// TIA Portal V20 export
VAR_GLOBAL   // PLC tag table "LASER_IN_datalogic"
   LASER_OFF AT %I400.0 : Bool;
   LASER_WARM_UP AT %I400.1 : Bool;
   LASER_WAIT_FOR_START AT %I400.2 : Bool;
   LASER_STANDBY AT %I400.3 : Bool;
   LASER_STANDBY_SHUTTER_CLOSED AT %I400.4 : Bool;
   LASER_READY AT %I400.5 : Bool;
   LASER_EMISSION AT %I400.6 : Bool;
   LASER_BUSSY_SHUTTER_CLOSED AT %I401.0 : Bool;
   LASER_WARNING AT %I401.1 : Bool;
   LASER_ERROR AT %I401.2 : Bool;
   COMMAND_EXECUTING AT %I402.0 : Bool;
   COMMAND_ERROR AT %I402.1 : Bool;
   PROTOCOL_ERROR AT %I402.2 : Bool;
   PROTOCOL_BOOT_UP AT %I403.7 : Bool;
   COMMAND_ERROR_CODE AT %IB404 : Byte;
   PROTOCOL_ERROR_CODE AT %IB405 : Byte;
   RESERVE_I_6_BYTE AT %IB406 : Byte;
   RESERVE_I_7_BYTE AT %IB407 : Byte;
   RESERVE_I_8_BYTE AT %IB408 : Byte;
   RESERVE_I_9_BYTE AT %IB409 : Byte;
   START_MARKING_IN AT %I410.0 : Bool;
   STOP_SYSTEM_IN AT %I410.1 : Bool;
   GET_PNIO_PROTOCOL_VERSION_IN AT %I411.0 : Bool;
   GET_LASER_ENGINE_VERSION AT %I411.1 : Bool;
   OPEN_DOCUMENT_FROM_DEVICE AT %I412.0 : Bool;
   SAVE_DOCUMENT AT %I412.1 : Bool;
   GET_DATA_FIELD_VALUE_IN AT %I412.2 : Bool;
   SET_DATA_FIELD_VALUE_IN AT %I412.3 : Bool;
   GET_GLOBAL_COUNTER_VALUE_IN AT %I412.4 : Bool;
   SET_GLOBAL_COUNTER_VALUE_IN AT %I412.5 : Bool;
   GET_GLOBAL_STRING_VALUE_IN AT %I412.6 : Bool;
   SET_GLOBAL_STRING_VALUE_IN AT %I412.7 : Bool;
   ENABLE_DATA_FIELD_IN AT %I413.0 : Bool;
   DISABLE_DATA_FIELD_IN AT %I413.1 : Bool;
   MOVE_END_ROTATE_DOCUMENT AT %I414.0 : Bool;
   MOVE_DATA_FIELD_IN AT %I414.1 : Bool;
   RESERVE_I_15_BYTE AT %IB415 : Byte;
   RESERVE_I_16_BYTE AT %IB416 : Byte;
   RESERVE_I_17_BYTE AT %IB417 : Byte;
   MOVE_AXIS_IN AT %I418.0 : Bool;
   RESET_AXIS_IN AT %I418.1 : Bool;
   STOP_AXIS_IN AT %I418.2 : Bool;
   START_AUTOFOCUS_IN AT %I418.3 : Bool;
   STOP_AUTOFOCUS_IN AT %I418.4 : Bool;
   SET_FOCUS_DISTANCE_REFERENCE_IN AT %I418.5 : Bool;
   RESERVE_I_19_BYTE AT %IB419 : Byte;
   X_AXIS_ENABLED AT %I420.0 : Bool;
   Y_AXIS_ENABLED AT %I420.1 : Bool;
   Z_AXIS_ENABLED AT %I420.2 : Bool;
   R_AXIS_ENABLED AT %I420.3 : Bool;
   X_AXIS_HOME AT %I420.4 : Bool;
   Y_AXIS_HOME AT %I420.5 : Bool;
   Z_AXIS_HOME AT %I420.6 : Bool;
   R_AXIS_HOME AT %I420.7 : Bool;
   X_AXIS_MOVEMENT AT %I421.0 : Bool;
   Y_AXIS_MOVEMENT AT %I421.1 : Bool;
   Z_AXIS_MOVEMENT AT %I421.2 : Bool;
   R_AXIS_MOVEMENT AT %I421.3 : Bool;
   Z_ASIS_IN_ON_FOCUS AT %I421.4 : Bool;
   FOCUS_DISTANCE_SENSOR_IS_AVAILABLE AT %I421.5 : Bool;
   RESERVE_I_22_BYTE AT %IB422 : Byte;
   RESERVE_I_23_BYTE AT %IB423 : Byte;
   SET_OUTPUT AT %I424.0 : Bool;
   RESET_OUTPUT_IN AT %I424.1 : Bool;
   RRESERVE_I_25_BYTE AT %IB425 : Byte;
   I_O_PORT_LASER_OUTPUT_STATUS_0 AT %I426.0 : Bool;
   I_O_PORT_LASER_OUTPUT_STATUS_1 AT %I426.1 : Bool;
   I_O_PORT_LASER_OUTPUT_STATUS_2 AT %I426.2 : Bool;
   I_O_PORT_LASER_OUTPUT_STATUS_3 AT %I426.3 : Bool;
   I_O_PORT_LASER_OUTPUT_STATUS_4 AT %I426.4 : Bool;
   I_O_PORT_LASER_OUTPUT_STATUS_5 AT %I426.5 : Bool;
   I_O_PORT_LASER_OUTPUT_STATUS_6 AT %I426.6 : Bool;
   I_O_PORT_LASER_OUTPUT_STATUS_7 AT %I426.7 : Bool;
   I_O_PORT_LASER_OUTPUT_STATUS_8 AT %I427.0 : Bool;
   I_O_PORT_LASER_OUTPUT_STATUS_9 AT %I427.1 : Bool;
   I_O_PORT_LASER_OUTPUT_STATUS_10 AT %I427.2 : Bool;
   I_O_PORT_LASER_OUTPUT_STATUS_11 AT %I427.3 : Bool;
   I_O_PORT_LASER_OUTPUT_STATUS_12 AT %I427.4 : Bool;
   I_O_PORT_LASER_OUTPUT_STATUS_13 AT %I427.5 : Bool;
   I_O_PORT_LASER_OUTPUT_STATUS_14 AT %I427.6 : Bool;
   I_O_PORT_LASER_OUTPUT_STATUS_15 AT %I427.7 : Bool;
   I_O_PORT_LASER_INPUT_STATUS_0 AT %I428.0 : Bool;
   I_O_PORT_LASER_INPUT_STATUS_1 AT %I428.1 : Bool;
   I_O_PORT_LASER_INPUT_STATUS_2 AT %I428.2 : Bool;
   I_O_PORT_LASER_INPUT_STATUS_3 AT %I428.3 : Bool;
   I_O_PORT_LASER_INPUT_STATUS_4 AT %I428.4 : Bool;
   I_O_PORT_LASER_INPUT_STATUS_5 AT %I428.5 : Bool;
   I_O_PORT_LASER_INPUT_STATUS_6 AT %I428.6 : Bool;
   I_O_PORT_LASER_INPUT_STATUS_7 AT %I428.7 : Bool;
   I_O_PORT_LASER_INPUT_STATUS_8 AT %I429.0 : Bool;
   I_O_PORT_LASER_INPUT_STATUS_9 AT %I429.1 : Bool;
   I_O_PORT_LASER_INPUT_STATUS_10 AT %I429.2 : Bool;
   I_O_PORT_LASER_INPUT_STATUS_11 AT %I429.3 : Bool;
   I_O_PORT_LASER_INPUT_STATUS_12 AT %I429.4 : Bool;
   I_O_PORT_LASER_INPUT_STATUS_13 AT %I429.5 : Bool;
   I_O_PORT_LASER_INPUT_STATUS_14 AT %I429.6 : Bool;
   I_O_PORT_LASER_INPUT_STATUS_15 AT %I429.7 : Bool;
   RESERVE_I_30_BYTE AT %IB430 : Byte;
   RESERVE_I_31_BYTE AT %IB431 : Byte;
   RESERVE_I_32_BYTE AT %IB432 : Byte;
   RESERVE_I_33_BYTE AT %IB433 : Byte;
   GET_ID_MATCH_RESULT_IN AT %I434.1 : Bool;
   GET_ID_MARVIS_CONFIGURATION_IN AT %I434.2 : Bool;
   SET_ID_MARVIS_CONFIGURATION_IN AT %I434.3 : Bool;
   GET_ID_MARVIS_RESULT_IN AT %I434.4 : Bool;
   RESERVE_I_35_BYTE AT %IB435 : Byte;
   MARVIS_RESULT_OK AT %I436.0 : Bool;
   MARVIS_RESULT_FAIL AT %I436.1 : Bool;
   SYMBOL_READ_OK AT %I436.2 : Bool;
   SYMBOL_READ_FAIL AT %I436.3 : Bool;
   SYMBOL_GRADE_RESULT_OK AT %I436.4 : Bool;
   SYMBOL_GRADE_RESULT_FAIL AT %I436.5 : Bool;
   SYMBOL_MATCH_RESULT_OK AT %I436.6 : Bool;
   SYMBOL_MATCH_RESULT_FAIL AT %I436.7 : Bool;
   RESERVE_I_37_BYTE AT %IB437 : Byte;
   READER_STATUS_AVAILABLE AT %I438.1 : Bool;
   READER_STATUS_BZSY AT %I438.2 : Bool;
   READER_STATUS_WARNING AT %I438.3 : Bool;
   READER_STATUS_ERROR AT %I438.4 : Bool;
   RESERVE_I_39_BYTE AT %IB439 : Byte;
   RESERVE_I_40_BYTE AT %IB440 : Byte;
   RESERVE_I_41_BYTE AT %IB441 : Byte;
   RESERVE_I_42_BYTE AT %IB442 : Byte;
   RESERVE_I_43_BYTE AT %IB443 : Byte;
   RESERVE_I_44_BYTE AT %IB444 : Byte;
   RESERVE_I_45_BYTE AT %IB445 : Byte;
   RESERVE_I_46_BYTE AT %IB446 : Byte;
   RESERVE_I_47_BYTE AT %IB447 : Byte;
   RESERVE_I_48_BYTE AT %IB448 : Byte;
   RESERVE_I_49_BYTE AT %IB449 : Byte;
   RESERVE_I_50_BYTE AT %IB450 : Byte;
   RESERVE_I_51_BYTE AT %IB451 : Byte;
   RESERVE_I_52_BYTE AT %IB452 : Byte;
   RESERVE_I_53_BYTE AT %IB453 : Byte;
   RESPONSE_DATE_SIZE AT %IB454 : Byte;
   RESERVE_I_55_BYTE AT %IB455 : Byte;
   RESPONSE_DATA_FIELD_0 AT %IB456 : Byte;
   RESPONSE_DATA_FIELD_1 AT %IB457 : Byte;
   RESPONSE_DATA_FIELD_2 AT %IB458 : Byte;
   RESPONSE_DATA_FIELD_3 AT %IB459 : Byte;
   RESPONSE_DATA_FIELD_4 AT %IB460 : Byte;
   RESPONSE_DATA_FIELD_5 AT %IB461 : Byte;
   RESPONSE_DATA_FIELD_6 AT %IB462 : Byte;
   RESPONSE_DATA_FIELD_7 AT %IB463 : Byte;
   RESPONSE_DATA_FIELD_8 AT %IB464 : Byte;
   RESPONSE_DATA_FIELD_9 AT %IB465 : Byte;
   RESPONSE_DATA_FIELD_10 AT %IB466 : Byte;
   RESPONSE_DATA_FIELD_11 AT %IB467 : Byte;
   RESPONSE_DATA_FIELD_12 AT %IB468 : Byte;
   RESPONSE_DATA_FIELD_13 AT %IB469 : Byte;
   RESPONSE_DATA_FIELD_14 AT %IB470 : Byte;
   RESPONSE_DATA_FIELD_15 AT %IB471 : Byte;
   RESPONSE_DATA_FIELD_16 AT %IB472 : Byte;
   RESPONSE_DATA_FIELD_17 AT %IB473 : Byte;
   RESPONSE_DATA_FIELD_18 AT %IB474 : Byte;
   RESPONSE_DATA_FIELD_19 AT %IB475 : Byte;
   RESPONSE_DATA_FIELD_20 AT %IB476 : Byte;
   RESPONSE_DATA_FIELD_21 AT %IB477 : Byte;
   RESPONSE_DATA_FIELD_22 AT %IB478 : Byte;
   RESPONSE_DATA_FIELD_23 AT %IB479 : Byte;
   RESPONSE_DATA_FIELD_24 AT %IB480 : Byte;
   RESPONSE_DATA_FIELD_25 AT %IB481 : Byte;
   RESPONSE_DATA_FIELD_26 AT %IB482 : Byte;
   RESPONSE_DATA_FIELD_27 AT %IB483 : Byte;
   RESPONSE_DATA_FIELD_28 AT %IB484 : Byte;
   RESPONSE_DATA_FIELD_29 AT %IB485 : Byte;
   RESPONSE_DATA_FIELD_30 AT %IB486 : Byte;
   RESPONSE_DATA_FIELD_31 AT %IB487 : Byte;
   RESPONSE_DATA_FIELD_32 AT %IB488 : Byte;
   RESPONSE_DATA_FIELD_33 AT %IB489 : Byte;
   RESPONSE_DATA_FIELD_34 AT %IB490 : Byte;
   RESPONSE_DATA_FIELD_35 AT %IB491 : Byte;
   RESPONSE_DATA_FIELD_36 AT %IB492 : Byte;
   RESPONSE_DATA_FIELD_37 AT %IB493 : Byte;
   RESPONSE_DATA_FIELD_38 AT %IB494 : Byte;
   RESPONSE_DATA_FIELD_39 AT %IB495 : Byte;
   RESPONSE_DATA_FIELD_40 AT %IB496 : Byte;
   RESPONSE_DATA_FIELD_41 AT %IB497 : Byte;
   RESPONSE_DATA_FIELD_42 AT %IB498 : Byte;
   RESPONSE_DATA_FIELD_43 AT %IB499 : Byte;
   RESPONSE_DATA_FIELD_44 AT %IB500 : Byte;
   RESPONSE_DATA_FIELD_45 AT %IB501 : Byte;
   RESPONSE_DATA_FIELD_46 AT %IB502 : Byte;
   RESPONSE_DATA_FIELD_47 AT %IB503 : Byte;
   RESPONSE_DATA_FIELD_48 AT %IB504 : Byte;
   RESPONSE_DATA_FIELD_49 AT %IB505 : Byte;
   RESPONSE_DATA_FIELD_50 AT %IB506 : Byte;
   RESPONSE_DATA_FIELD_51 AT %IB507 : Byte;
   RESPONSE_DATA_FIELD_52 AT %IB508 : Byte;
   RESPONSE_DATA_FIELD_53 AT %IB509 : Byte;
   RESPONSE_DATA_FIELD_54 AT %IB510 : Byte;
   RESPONSE_DATA_FIELD_55 AT %IB511 : Byte;
   RESPONSE_DATA_FIELD_56 AT %IB512 : Byte;
   RESPONSE_DATA_FIELD_57 AT %IB513 : Byte;
   RESPONSE_DATA_FIELD_58 AT %IB514 : Byte;
   RESPONSE_DATA_FIELD_59 AT %IB515 : Byte;
   RESPONSE_DATA_FIELD_60 AT %IB516 : Byte;
   RESPONSE_DATA_FIELD_61 AT %IB517 : Byte;
   RESPONSE_DATA_FIELD_62 AT %IB518 : Byte;
   RESPONSE_DATA_FIELD_63 AT %IB519 : Byte;
   RESPONSE_DATA_FIELD_64 AT %IB520 : Byte;
   RESPONSE_DATA_FIELD_65 AT %IB521 : Byte;
   RESPONSE_DATA_FIELD_66 AT %IB522 : Byte;
   RESPONSE_DATA_FIELD_67 AT %IB523 : Byte;
   RESPONSE_DATA_FIELD_68 AT %IB524 : Byte;
   RESPONSE_DATA_FIELD_69 AT %IB525 : Byte;
   RESPONSE_DATA_FIELD_70 AT %IB526 : Byte;
   RESPONSE_DATA_FIELD_71 AT %IB527 : Byte;
END_VAR
